(* IEC 61131-3 sources: rusty/tests/lit/multi/polymorphism_class, 5 files *)

(* ---- main.st ---- *)
FUNCTION main
    VAR
        instanceA: ClassA;
        instanceB: ClassB;
        instanceC: ClassC;
        instanceD: ClassD;

        refInstanceA: POINTER TO ClassA;
    END_VAR

    refInstanceA := ADR(instanceA);
    refInstanceA^.alpha();
    refInstanceA^.bravo();
    refInstanceA^.charlie();
    refInstanceA^.delta();

    refInstanceA := ADR(instanceB);
    refInstanceA^.alpha();
    refInstanceA^.bravo();
    refInstanceA^.charlie();
    refInstanceA^.delta();

    refInstanceA := ADR(instanceC);
    refInstanceA^.alpha();
    refInstanceA^.bravo();
    refInstanceA^.charlie();
    refInstanceA^.delta();

    refInstanceA := ADR(instanceD);
    refInstanceA^.alpha();
    refInstanceA^.bravo();
    refInstanceA^.charlie();
    refInstanceA^.delta();
END_FUNCTION

(* ---- a.st ---- *)
CLASS ClassA
    METHOD alpha
        printf('ClassA::alpha$N');
    END_METHOD

    METHOD bravo
        printf('ClassA::bravo$N');
    END_METHOD

    METHOD charlie
        printf('ClassA::charlie$N');
    END_METHOD

    METHOD delta
        printf('ClassA::delta$N');
    END_METHOD
END_CLASS

(* ---- b.st ---- *)
CLASS ClassB EXTENDS ClassA
    METHOD bravo
        printf('ClassB::bravo$N');
    END_METHOD
END_CLASS

(* ---- c.st ---- *)
CLASS ClassC EXTENDS ClassB
    METHOD charlie
        printf('ClassC::charlie$N');
    END_METHOD
END_CLASS

(* ---- d.st ---- *)
CLASS ClassD EXTENDS ClassC
    METHOD alpha
        printf('ClassD::alpha$N');
    END_METHOD

    METHOD bravo
        printf('ClassD::bravo$N');
    END_METHOD

    METHOD charlie
        printf('ClassD::charlie$N');
    END_METHOD

    METHOD delta
        printf('ClassD::delta$N');
    END_METHOD
END_CLASS
